Fanuc KAREL source: KO00009.KL

PROGRAM KO00009
%NOLOCKGROUP
VAR
  P1: XYZWPR
  P2: XYZWPR
  P3: XYZWPR
  OUT: POSITION
BEGIN
  OUT = FRAME(P1, P2, P3)
END KO00009
